// Generated by voz_llm_plc_agent
// Target: Siemens TIA Portal V18 - SCL external source
// Review and compile before any download to physical hardware.

FUNCTION_BLOCK "PLC_PRG"
{ S7_Optimized_Access := 'TRUE' }
VERSION : 0.1
VAR_INPUT
   I_Start : Bool := FALSE;
   I_Emergency : Bool := FALSE;
END_VAR
VAR_OUTPUT
   Q_Motor_Enable : Bool := FALSE;
END_VAR
VAR
   M_RunLatch : Bool;
   T_OperationLimit {InstructionName := 'TON_TIME'; LibVersion := '1.0'} : TON_TIME;
   M_Motor_EnableLatch : Bool;
END_VAR
BEGIN
(* Paro automatico del motor por tiempo de operacion *)
IF #I_Emergency OR FALSE THEN
    #M_RunLatch := FALSE;
ELSIF #I_Start THEN
    #M_RunLatch := TRUE;
END_IF;

#T_OperationLimit(IN := #M_RunLatch AND NOT #I_Emergency, PT := T#10s);

IF #T_OperationLimit.Q THEN
    #M_RunLatch := FALSE;
END_IF;

#Q_Motor_Enable := #M_RunLatch AND NOT #I_Emergency;
END_FUNCTION_BLOCK

DATA_BLOCK "DB_PLC_PRG"
{ S7_Optimized_Access := 'TRUE' }
VERSION : 0.1
NON_RETAIN
"PLC_PRG"
BEGIN
END_DATA_BLOCK

ORGANIZATION_BLOCK "Main"
{ S7_Optimized_Access := 'TRUE' }
VERSION : 0.1
BEGIN
   "DB_PLC_PRG"(
      I_Start := "I_Start",
      I_Emergency := "I_Emergency",
      Q_Motor_Enable => "Q_Motor_Enable"
   );
END_ORGANIZATION_BLOCK
